FUNCTION_BLOCK "fb_bancoEt200_32"
TITLE = fb_bancoEt200_32 v0.1
{ S7_Optimized_Access := 'TRUE' }
AUTHOR : 'RegLobo'
VERSION : 0.1
////====================================
//// fb_bancoEt200_32  -  RASCUNHO v0.1 (03/11/2026) GERADO por gerar_banco_v0.2.py - nao compilado, nao testado
//// ONDE RODA : ET200 (programa Gerador_BC015). 1 instancia por banco NOVO (BC550, BC59,5). BC56 e BC400 seguem no FC4 atual.
//// O QUE FAZ : lado ET200 do telegrama PUT/GET do banco (ate 32 chaves, 8+8 bytes):
////    1) vidaET incrementa a cada ~100 ms (prova ao 1515 que o ET200 esta vivo).
////    2) vida1515 parou de mudar por TempoPerdaMs -> ComOk=FALSE e TODAS as saidas vao a FALSE.
////    3) apos queda, a chave so religa depois de o comando cair a FALSE e ser recomandado (nao religa sozinha).
////    4) saida da contatora so liga com ComOk E LigarBanco E seletora em Auto (defesa extra; o 1515 ja zera o comando).
////    5) fbk[n] = contato auxiliar REAL; seletoraAuto = entrada fisica da seletora do banco (1 = Auto).
//// COMO CHAMAR: ver fc_bancosNovosEt200 (gerado). Entradas/saidas fisicas entram pelas tags da tabela tags_ET200_bancos.
////=====================================
   VAR_INPUT
      NumChaves        : Int;                       // chaves reais deste banco (1..32)
      SeletoraEntrada  : Bool;                      // entrada fisica: seletora do banco em Auto (1 = Auto)
      TempoPerdaMs     : Time := T#2S;              // menor que o TempoVida do 1515 (3 s)
   END_VAR
   VAR_OUTPUT
      ComOk : Bool;
   END_VAR
   VAR_IN_OUT
      Cmd               : Array[1..32] of Bool;   // <DB remoto>.cmd       (PUT do 1515; so le)
      Vida1515          : Int;                     // <DB remoto>.vida1515  (so le)
      LigarBanco        : Bool;                    // <DB remoto>.ligarBanco (so le)
      VidaET            : Int;                     // <DB remoto>.vidaET    (escreve)
      Fbk               : Array[1..32] of Bool;   // <DB remoto>.fbk       (escreve)
      SeletoraAuto      : Bool;                    // <DB remoto>.seletoraAuto (escreve)
      SaidaContatora    : Array[1..32] of Bool;   // saidas fisicas (copiadas pelo fc_bancosNovosEt200)
      EntradaContatoAux : Array[1..32] of Bool;   // contatos auxiliares fisicos
   END_VAR
   VAR
      _tOsc100ms   : TON_TIME;
      _tPerda      : TON_TIME;
      _vida1515Ant : Int;
      _vidaMudou   : Bool;
      _comOkAnt    : Bool;
      _cmdAnt      : Array[1..32] of Bool;
      _rearmado    : Array[1..32] of Bool;
      i            : Int;
   END_VAR

BEGIN
   #_tOsc100ms(IN := NOT #_tOsc100ms.Q, PT := T#100MS);
   IF #_tOsc100ms.Q THEN
      #VidaET := #VidaET + 1;
      IF #VidaET >= 32767 THEN #VidaET := 0; END_IF;
   END_IF;

   IF #Vida1515 <> #_vida1515Ant THEN
      #_vida1515Ant := #Vida1515;
      #_vidaMudou := TRUE;
   ELSE
      #_vidaMudou := FALSE;
   END_IF;
   #_tPerda(IN := NOT #_vidaMudou, PT := #TempoPerdaMs);   // vida nova reseta; sem vida nova conta
   #ComOk := NOT #_tPerda.Q;

   IF #ComOk AND NOT #_comOkAnt THEN
      FOR #i := 1 TO #NumChaves DO
         #_rearmado[#i] := FALSE;
      END_FOR;
   END_IF;

   #SeletoraAuto := #SeletoraEntrada;

   FOR #i := 1 TO 32 DO
      IF #i <= #NumChaves THEN
         #Fbk[#i] := #EntradaContatoAux[#i];
         IF NOT #Cmd[#i] AND #_cmdAnt[#i] THEN
            #_rearmado[#i] := TRUE;
         END_IF;
         IF #ComOk AND #LigarBanco AND #SeletoraEntrada AND (#_comOkAnt OR #_rearmado[#i]) THEN
            #SaidaContatora[#i] := #Cmd[#i];
         ELSE
            #SaidaContatora[#i] := FALSE;
         END_IF;
         #_cmdAnt[#i] := #Cmd[#i];
      ELSE
         #Fbk[#i] := FALSE;
         #SaidaContatora[#i] := FALSE;
      END_IF;
   END_FOR;

   #_comOkAnt := #ComOk;
END_FUNCTION_BLOCK
